TYPE U_YARD_STATE :
UNION
  stState             : ST_YARD_STATE;
  byState   AT %Q*    : ARRAY[1..SIZEOF(ST_YARD_STATE)] OF BYTE;
END_UNION
END_TYPE

(* stored: Version 1.1.0.1
   DUT U_YARD_STATE: Id {420ba58f-f9f5-4337-9e40-e89ae279ac58} *)
